Staubli VAL3: Algorithm6.dtx

public num nInverseMatrix1[4 4]
  [0,0] = 1.945193
  [0,1] = -1.712762
  [0,2] = 9.261268
  [1,0] = 0.502721
  [1,1] = 0.619141
  [1,2] = -1.663322
  [2,0] = 0.453432
  [2,1] = 1.0601144
  [2,2] = 3.220251
  [3,3] = 1
public num nMatrix1[4 4]
  [0,0] = 0.27407
  [0,1] = 1.118537
  [0,2] = -0.210464
  [1,0] = -0.17311
  [1,1] = 0.150611
  [1,2] = 0.575649
  [2,0] = 0.0183975
  [2,1] = -0.207079
  [2,2] = 0.150664
  [3,3] = 1
public num nMatrix2[4 4]
  [0,0] = 1
  [1,1] = 1
  [2,2] = 1
  [3,0] = 31.552388
  [3,1] = 103.369183
  [3,2] = -8.232965
  [3,3] = 1
public num nMatrix3[4 4]
  [0,0] = 1.945193
  [0,1] = -1.712762
  [0,2] = 9.261268
  [1,0] = 0.502721
  [1,1] = 0.619141
  [1,2] = -1.663322
  [2,0] = 0.453432
  [2,1] = 1.0601144
  [2,2] = 3.220251
  [3,0] = 109.608277
  [3,1] = 1.230419
  [3,2] = 93.766659
  [3,3] = 1
public num nTeach_3_1[4 4]
  [0,0] = -0.024705
  [0,1] = -0.0184623
  [0,2] = -0.999524
  [1,0] = -0.240476
  [1,1] = 0.970581
  [1,2] = -0.0119839
  [2,0] = 0.970341
  [2,1] = 0.240066
  [2,2] = -0.028418
  [3,0] = 888.833618
  [3,1] = -160.122184
  [3,2] = -41.507861
  [3,3] = 1
public num nTeach_3_2[4 4]
  [0,0] = -0.298775
  [0,1] = 0.518277
  [0,2] = -0.801326
  [1,0] = -0.0673661
  [1,1] = 0.82613
  [1,2] = 0.559438
  [2,0] = 0.951943
  [2,1] = 0.221128
  [2,2] = -0.211913
  [3,0] = 920.386007
  [3,1] = -217.720531
  [3,2] = -46.252531
  [3,3] = 1
public num nTeach_3_3[4 4]
  [0,0] = 0.130655
  [0,1] = -0.60026
  [0,2] = -0.789061
  [1,0] = -0.445377
  [1,1] = 0.67552
  [1,2] = -0.587633
  [2,0] = 0.885759
  [2,1] = 0.428207
  [2,2] = -0.179082
  [3,0] = 879.830904
  [3,1] = -114.351348
  [3,2] = -49.740826
  [3,3] = 1
